(* LS Electric XG5000 project: NewProject *)
(* PLC LSPLC *)

FUNCTION UserDouble : DINT
(* Doubles an integer *)
VAR_INPUT
    Value : DINT;
END_VAR
UserDouble := Value * 2;
END_FUNCTION

FUNCTION_BLOCK UserAccumulator
(* State retained by each instance between calls *)
VAR_INPUT
    Reset : BOOL;
    Increment : DINT;
END_VAR
VAR_OUTPUT
    Total : DINT;
END_VAR
IF Reset THEN
    Total := 0;
ELSE
    Total := Total + Increment;
END_IF;
END_FUNCTION_BLOCK

FUNCTION UserCopyBOOL : BOOL
VAR_INPUT
    Value : BOOL;
    Second : BOOL;
END_VAR
VAR_IN_OUT
    Shared : BOOL;
END_VAR
UserCopyBOOL := Value;
END_FUNCTION

FUNCTION UserCopyBYTE : BYTE
VAR_INPUT
    Value : BYTE;
    Second : BYTE;
END_VAR
VAR_IN_OUT
    Shared : BYTE;
END_VAR
UserCopyBYTE := Value;
END_FUNCTION

FUNCTION UserCopyWORD : WORD
VAR_INPUT
    Value : WORD;
    Second : WORD;
END_VAR
VAR_IN_OUT
    Shared : WORD;
END_VAR
UserCopyWORD := Value;
END_FUNCTION

FUNCTION UserCopyDWORD : DWORD
VAR_INPUT
    Value : DWORD;
    Second : DWORD;
END_VAR
VAR_IN_OUT
    Shared : DWORD;
END_VAR
UserCopyDWORD := Value;
END_FUNCTION

FUNCTION UserCopyLWORD : LWORD
VAR_INPUT
    Value : LWORD;
    Second : LWORD;
END_VAR
VAR_IN_OUT
    Shared : LWORD;
END_VAR
UserCopyLWORD := Value;
END_FUNCTION

FUNCTION UserCopySINT : SINT
VAR_INPUT
    Value : SINT;
    Second : SINT;
END_VAR
VAR_IN_OUT
    Shared : SINT;
END_VAR
UserCopySINT := Value;
END_FUNCTION

FUNCTION UserCopyINT : INT
VAR_INPUT
    Value : INT;
    Second : INT;
END_VAR
VAR_IN_OUT
    Shared : INT;
END_VAR
UserCopyINT := Value;
END_FUNCTION

FUNCTION UserCopyDINT : DINT
VAR_INPUT
    Value : DINT;
    Second : DINT;
END_VAR
VAR_IN_OUT
    Shared : DINT;
END_VAR
UserCopyDINT := Value;
END_FUNCTION

FUNCTION UserCopyLINT : LINT
VAR_INPUT
    Value : LINT;
    Second : LINT;
END_VAR
VAR_IN_OUT
    Shared : LINT;
END_VAR
UserCopyLINT := Value;
END_FUNCTION

FUNCTION UserCopyUSINT : USINT
VAR_INPUT
    Value : USINT;
    Second : USINT;
END_VAR
VAR_IN_OUT
    Shared : USINT;
END_VAR
UserCopyUSINT := Value;
END_FUNCTION

FUNCTION UserCopyUINT : UINT
VAR_INPUT
    Value : UINT;
    Second : UINT;
END_VAR
VAR_IN_OUT
    Shared : UINT;
END_VAR
UserCopyUINT := Value;
END_FUNCTION

FUNCTION UserCopyUDINT : UDINT
VAR_INPUT
    Value : UDINT;
    Second : UDINT;
END_VAR
VAR_IN_OUT
    Shared : UDINT;
END_VAR
UserCopyUDINT := Value;
END_FUNCTION

FUNCTION UserCopyULINT : ULINT
VAR_INPUT
    Value : ULINT;
    Second : ULINT;
END_VAR
VAR_IN_OUT
    Shared : ULINT;
END_VAR
UserCopyULINT := Value;
END_FUNCTION

FUNCTION UserCopyREAL : REAL
VAR_INPUT
    Value : REAL;
    Second : REAL;
END_VAR
VAR_IN_OUT
    Shared : REAL;
END_VAR
UserCopyREAL := Value;
END_FUNCTION

FUNCTION UserCopyLREAL : LREAL
VAR_INPUT
    Value : LREAL;
    Second : LREAL;
END_VAR
VAR_IN_OUT
    Shared : LREAL;
END_VAR
UserCopyLREAL := Value;
END_FUNCTION

FUNCTION UserCopyTIME : TIME
VAR_INPUT
    Value : TIME;
    Second : TIME;
END_VAR
VAR_IN_OUT
    Shared : TIME;
END_VAR
UserCopyTIME := Value;
END_FUNCTION

FUNCTION UserCopyDATE : DATE
VAR_INPUT
    Value : DATE;
    Second : DATE;
END_VAR
VAR_IN_OUT
    Shared : DATE;
END_VAR
UserCopyDATE := Value;
END_FUNCTION

FUNCTION UserCopyTIME_OF_DAY : TIME_OF_DAY
VAR_INPUT
    Value : TIME_OF_DAY;
    Second : TIME_OF_DAY;
END_VAR
VAR_IN_OUT
    Shared : TIME_OF_DAY;
END_VAR
UserCopyTIME_OF_DAY := Value;
END_FUNCTION

FUNCTION UserCopyDATE_AND_TIME : DATE_AND_TIME
VAR_INPUT
    Value : DATE_AND_TIME;
    Second : DATE_AND_TIME;
END_VAR
VAR_IN_OUT
    Shared : DATE_AND_TIME;
END_VAR
UserCopyDATE_AND_TIME := Value;
END_FUNCTION

FUNCTION_BLOCK UserAllScalars
VAR_INPUT
    ValueBOOL : BOOL;
    ValueBYTE : BYTE;
    ValueWORD : WORD;
    ValueDWORD : DWORD;
    ValueLWORD : LWORD;
    ValueSINT : SINT;
    ValueINT : INT;
    ValueDINT : DINT;
    ValueLINT : LINT;
    ValueUSINT : USINT;
    ValueUINT : UINT;
    ValueUDINT : UDINT;
    ValueULINT : ULINT;
    ValueREAL : REAL;
    ValueLREAL : LREAL;
    ValueTIME : TIME;
    ValueDATE : DATE;
    ValueTIME_OF_DAY : TIME_OF_DAY;
    ValueDATE_AND_TIME : DATE_AND_TIME;
    ExtraBool : BOOL;
END_VAR
VAR_IN_OUT
    SharedBOOL : BOOL;
    SharedBYTE : BYTE;
    SharedWORD : WORD;
    SharedDWORD : DWORD;
    SharedLWORD : LWORD;
    SharedSINT : SINT;
    SharedINT : INT;
    SharedDINT : DINT;
    SharedLINT : LINT;
    SharedUSINT : USINT;
    SharedUINT : UINT;
    SharedUDINT : UDINT;
    SharedULINT : ULINT;
    SharedREAL : REAL;
    SharedLREAL : LREAL;
    SharedTIME : TIME;
    SharedDATE : DATE;
    SharedTIME_OF_DAY : TIME_OF_DAY;
    SharedDATE_AND_TIME : DATE_AND_TIME;
END_VAR
VAR_OUTPUT
    OutputBOOL : BOOL;
    OutputBYTE : BYTE;
    OutputWORD : WORD;
    OutputDWORD : DWORD;
    OutputLWORD : LWORD;
    OutputSINT : SINT;
    OutputINT : INT;
    OutputDINT : DINT;
    OutputLINT : LINT;
    OutputUSINT : USINT;
    OutputUINT : UINT;
    OutputUDINT : UDINT;
    OutputULINT : ULINT;
    OutputREAL : REAL;
    OutputLREAL : LREAL;
    OutputTIME : TIME;
    OutputDATE : DATE;
    OutputTIME_OF_DAY : TIME_OF_DAY;
    OutputDATE_AND_TIME : DATE_AND_TIME;
    Out : BOOL;
END_VAR
VAR
    Private : INT;
END_VAR
Private := 1;
Out := ValueBOOL;
END_FUNCTION_BLOCK

PROGRAM NewProgram (* task: 스캔 프로그램 *)
VAR
    Counter : UserAccumulator;
    Observed : DINT;
    Result : DINT;
END_VAR
Result := UserDouble(Value := 4);
Counter(Reset := FALSE, Increment := Result);
Observed := Counter.Total;
END_PROGRAM